SUBAPPLICATION AX_TO_QXA_BG_PUBLISH_SWITCHPIC_OPT (* Wie AX_TO_QXA_BG_PUBLISH_SWITCHPIC, aber mit 2 AOption-Sockets: AOption_Output schaltet nur den physischen Ausgang, AOption_Anzeige Hintergrund+Publish+ObjectPointer. INIT_CNF je echt zurueck. *)
  (* Standard: 61499-2; Description: Copyright (c) 2026 Meisterschulen am Ostbahnhof This program and the accompanying materials are made available under the terms of the Eclipse Public License 2.0 which is available at https://www.eclipse.org/legal/epl-2.0/ SPDX-License-Identifier: EPL-2.0 *)
  (* Version 1.0, 2026-10-16, Franz Höpfinger, Meisterschulen am Ostbahnhof, Kopie von AX_TO_QXA_BG_PUBLISH_SWITCHPIC v1.2 (Franz: 'Die Lib Typen KOPIEREN und die Kopie aendern') - statt QI/INIT 2 AOption-Sockets: AOption_Output (nur physischer Ausgang) und AOption_Anzeige (Hintergrund/Publish/ObjPtr). Grund: bei Igel/Elevator=PVEA blieben SoftKey-Hintergrund, ObjectPointer und State-Publish tot. *)
  PACKAGE MyLib::sys;
  IMPORT isobus::UT::Q::const::IDs::ID_NULL;
  IMPORT logiBUS::io::DQ::logiBUS_DO;
  IMPORT logiBUS::io::DQ::logiBUS_DO_S;
  IMPORT isobus::UT::Q::types::s2x1ObjectIDs;
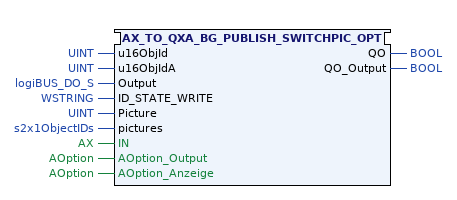
  VAR_INPUT
    u16ObjId : UINT := ID_NULL; (* Object ID Softkey - traegt die Hintergrundfarbe *)
    u16ObjIdA : UINT := ID_NULL; (* Object ID AuxFunction2 (Joystick) - zeigt Hintergrundfarbe am Aux-Handle mit *)
    Output : logiBUS::io::DQ::logiBUS_DO_S := logiBUS_DO::Invalid; (* Identify the Output Output_Q1..Q12 *)
    ID_STATE_WRITE : WSTRING; (* Lokale Publish-Adresse (ACTION=WRITE) fuer den Zustand - wird von Web-Client/Dashboard remote abonniert *)
    Picture : UINT; (* Object ID des ObjectPointer, der den Status-Kaestchen-Inhalt traegt *)
    pictures : isobus::UT::Q::types::s2x1ObjectIDs := (up := (u16ObjId := ID_NULL), down := (u16ObjId := ID_NULL)); (* die beiden Ziel-Object-IDs (up=aus, down=an) *)
  END_VAR
  VAR_OUTPUT
    QO : BOOL; (* Quality Output Anzeige (AND aus Publish/ObjPtr) *)
    QO_Output : BOOL; (* Quality Output physischer Ausgang *)
  END_VAR
  SOCKETS
    IN : adapter::types::unidirectional::AX; (* Fertiger AX-Zustand - wird auf Ausgang+Hintergrund+Publish UND ObjectPointer-Statusanzeige verteilt *)
    AOption_Output : Option::AOption; (* Aktiviert nur den physischen Ausgang (z.B. DEMUX-Zweig Klassisch) *)
    AOption_Anzeige : Option::AOption; (* Aktiviert Hintergrund+Publish+ObjectPointer (z.B. AOption_OR_2 aus Klassisch+PVEA) *)
  END_SOCKETS
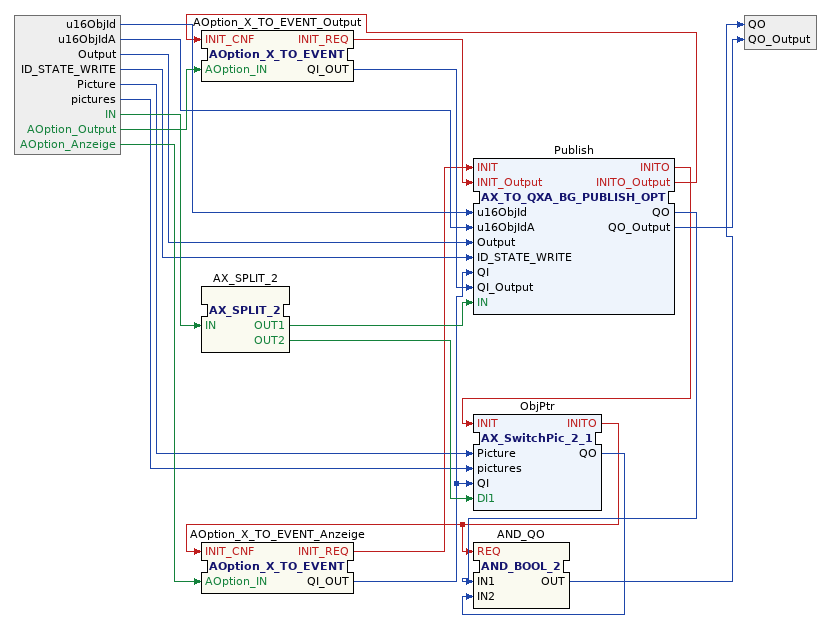
  FBS
    AX_SPLIT_2 : adapter::events::unidirectional::AX_SPLIT_2;
    AOption_X_TO_EVENT_Output : Option::conversion::AOption_X_TO_EVENT;
    AOption_X_TO_EVENT_Anzeige : Option::conversion::AOption_X_TO_EVENT;
    AND_QO : iec61131::booleanOperators::AND_BOOL_2;
  END_FBS
  SUBAPPS
    Publish : MyLib::sys::AX_TO_QXA_BG_PUBLISH_OPT;
    ObjPtr : MyLib::sys::AX_SwitchPic_2_1;
  END_SUBAPPS
  EVENT_CONNECTIONS
    AOption_X_TO_EVENT_Anzeige.INIT_REQ TO Publish.INIT;
    Publish.INITO TO ObjPtr.INIT;
    ObjPtr.INITO TO AND_QO.REQ;
    ObjPtr.INITO TO AOption_X_TO_EVENT_Anzeige.INIT_CNF;
    AOption_X_TO_EVENT_Output.INIT_REQ TO Publish.INIT_Output;
    Publish.INITO_Output TO AOption_X_TO_EVENT_Output.INIT_CNF;
  END_CONNECTIONS
  DATA_CONNECTIONS
    u16ObjId TO Publish.u16ObjId;
    u16ObjIdA TO Publish.u16ObjIdA;
    Output TO Publish.Output;
    ID_STATE_WRITE TO Publish.ID_STATE_WRITE;
    Picture TO ObjPtr.Picture;
    pictures TO ObjPtr.pictures;
    AOption_X_TO_EVENT_Anzeige.QI_OUT TO Publish.QI;
    AOption_X_TO_EVENT_Anzeige.QI_OUT TO ObjPtr.QI;
    AOption_X_TO_EVENT_Output.QI_OUT TO Publish.QI_Output;
    Publish.QO TO AND_QO.IN1;
    ObjPtr.QO TO AND_QO.IN2;
    AND_QO.OUT TO QO;
    Publish.QO_Output TO QO_Output;
  END_CONNECTIONS
  ADAPTER_CONNECTIONS
    IN TO AX_SPLIT_2.IN;
    AX_SPLIT_2.OUT1 TO Publish.IN;
    AX_SPLIT_2.OUT2 TO ObjPtr.DI1;
    AOption_Output TO AOption_X_TO_EVENT_Output.AOption_IN;
    AOption_Anzeige TO AOption_X_TO_EVENT_Anzeige.AOption_IN;
  END_CONNECTIONS
END_SUBAPPLICATION
